INTERFACE I_FillValve EXTENDS I_Diagnosable

METHOD Open
END_METHOD

METHOD Close
END_METHOD

PROPERTY IsOpen : BOOL
GET
END_GET
END_PROPERTY

PROPERTY IsClosed : BOOL
GET
END_GET
END_PROPERTY

END_INTERFACE

(* stored: Version 1.1.0.1
   Itf I_FillValve: Id {6afaa988-396f-4c42-8a97-f9acf02797c2}
   Method Open: Id {da2bbfd5-35f4-49e0-9d55-92f89caa1fc8}
   Method Close: Id {4bfd4cfa-1844-48a5-8f63-1a336ab2f40f}
   Property IsOpen: Id {727a8224-d15f-4d6f-900e-b1d96dc0f499}
   Get Get: Id {05232500-5fb4-4dd3-a509-f963d50b260d}
   Property IsClosed: Id {3460cd2c-b32d-46f0-a8bd-cda99bc392a6}
   Get Get: Id {85f84552-2f09-410d-b45d-6e2cf4a62259} *)
